TYPE EthercatDevice :
STRUCT
	mDirection AT %Q*: BOOL ;
	mSpeed AT %Q*: DWORD ;
	mTime AT %Q*: DWORD ;
	mMode AT %Q*: BOOL ;
END_STRUCT
END_TYPE

(* stored: Version 1.1.0.1, ProductVersion 3.1.4024.11
   DUT EthercatDevice: Id {b0ed898d-e1ad-436f-8e91-59112c261c39} *)
